(* IEC 61131-3 sources: Jacob-Formschaumtechnik-ISEL-CNC-Retrofit/twincat/PLC/src/5_Messages, 3 files *)

(* ---- F_ToFaultClass.st ---- *)
FUNCTION F_ToFaultClass : E_FaultClass
VAR_INPUT
    nClass : INT;
END_VAR

CASE nClass OF
    0: F_ToFaultClass := E_FaultClass.R0_Info;
    1: F_ToFaultClass := E_FaultClass.R1_Warning;
    2: F_ToFaultClass := E_FaultClass.R2_FeedHold;
    3: F_ToFaultClass := E_FaultClass.R3_Abort;
ELSE
    F_ToFaultClass := E_FaultClass.R4_DrivesOff;   (* unbekannt: sicherste Reaktion *)
END_CASE
END_FUNCTION

(* ---- FB_AlarmJournal.st ---- *)
(* Meldejournal (Anforderung 2.9.2, Befund 21): Ringpuffer der letzten 100 kommenden Meldungen
   mit Klasse und Zeitstempel (UTC aus F_GetSystemTime). Ablage in GVL_Persistent.stJournal,
   die HMI liest die Kopie GVL_HMI.stJournal. Spaeter optional zusaetzlich Tc3_EventLogger. *)
FUNCTION_BLOCK FB_AlarmJournal
VAR_INPUT
    aCond : ARRAY[0..14] OF BOOL;
    aId   : ARRAY[0..14] OF INT;
    aClass: ARRAY[0..14] OF INT;
    dtNow : DT;
END_VAR
VAR_IN_OUT
    stJournal : ST_HmiJournal;
END_VAR
VAR_OUTPUT
    nEntries : UINT;
    bChanged : BOOL;      (* in diesem Zyklus neuer Eintrag *)
END_VAR
VAR
    aPrev  : ARRAY[0..14] OF BOOL;
    i      : INT;
END_VAR

bChanged := FALSE;
IF stJournal.nHead > 99 THEN stJournal.nHead := 0; END_IF   (* Schutz bei beschaedigten Persistenzdaten *)
FOR i := 0 TO 14 DO
    IF aCond[i] AND NOT aPrev[i] THEN
        stJournal.aEntry[stJournal.nHead].nId    := aId[i];
        stJournal.aEntry[stJournal.nHead].nClass := aClass[i];
        stJournal.aEntry[stJournal.nHead].dtTime := dtNow;
        stJournal.nHead := (stJournal.nHead + 1) MOD 100;
        IF stJournal.nEntries < 100 THEN stJournal.nEntries := stJournal.nEntries + 1; END_IF
        stJournal.nSeq := stJournal.nSeq + 1;
        bChanged := TRUE;
    END_IF
    aPrev[i] := aCond[i];
END_FOR
nEntries := stJournal.nEntries;
END_FUNCTION_BLOCK

(* ---- FB_AlarmList.st ---- *)
(* Zentrale Meldeliste. Die Logik setzt aCond[Slot] jeden Zyklus, solange die Ursache besteht.
   R3 und R4 bleiben nach Wegfall der Ursache gespeichert, bis quittiert wird (Wiederanlauf nie
   automatisch). Hoechste Klasse gewinnt, bei gleicher Klasse die kleinste ID.
   Anzeige an die HMI spaeter ueber Tc3_EventLogger (Adapter), die Logik bleibt unabhaengig. *)
FUNCTION_BLOCK FB_AlarmList
VAR_INPUT
    aCond : ARRAY[0..14] OF BOOL;        (* Index = E_AlarmSlot *)
    bAck  : BOOL;                        (* Impuls: gespeicherte Meldungen quittieren *)
END_VAR
VAR_OUTPUT
    nActive        : UINT;
    nTopId         : INT;
    nTopClass      : INT;                (* 0..4 = E_FaultClass, Umwandlung mit F_ToFaultClass *)
    bAnyR2OrHigher : BOOL;
    bAnyR3OrHigher : BOOL;
    bAnyR4         : BOOL;
    bAckPending    : BOOL;               (* gespeicherte R3/R4 warten auf Quittierung *)
    aList          : ARRAY[0..14] OF ST_Alarm;   (* fuer die HMI *)
END_VAR
VAR
    aId    : ARRAY[0..14] OF INT;      (* Kopie aus GVL_AlarmCatalog *)
    aClass : ARRAY[0..14] OF INT;
    aLatch : ARRAY[0..14] OF BOOL;
    i      : INT;
    rtAck  : R_TRIG;
    nCls   : INT;
END_VAR

aId := GVL_AlarmCatalog.aAlarmId;
aClass := GVL_AlarmCatalog.aAlarmClass;
rtAck(CLK := bAck);
nActive := 0; nTopId := 0; nTopClass := 0;
bAnyR2OrHigher := FALSE; bAnyR3OrHigher := FALSE; bAnyR4 := FALSE; bAckPending := FALSE;

FOR i := 0 TO 14 DO
    nCls := aClass[i];
    IF aCond[i] AND nCls >= 3 THEN
        aLatch[i] := TRUE;
    END_IF
    IF rtAck.Q AND NOT aCond[i] THEN
        aLatch[i] := FALSE;
    END_IF
    aList[i].nId := aId[i];
    aList[i].eClass := F_ToFaultClass(nCls);
    aList[i].bActive := aCond[i];
    aList[i].bLatched := aLatch[i] AND NOT aCond[i];
    IF aCond[i] OR aLatch[i] THEN
        nActive := nActive + 1;
        IF nCls >= 2 THEN bAnyR2OrHigher := TRUE; END_IF
        IF nCls >= 3 THEN bAnyR3OrHigher := TRUE; END_IF
        IF nCls = 4  THEN bAnyR4 := TRUE; END_IF
        IF aLatch[i] AND NOT aCond[i] THEN bAckPending := TRUE; END_IF
        IF nTopId = 0 OR nCls > nTopClass OR (nCls = nTopClass AND aId[i] < nTopId) THEN
            nTopId := aId[i];
            nTopClass := nCls;
        END_IF
    END_IF
END_FOR
END_FUNCTION_BLOCK
